(* IEC 61131-3 sources: kns-pump-station/src/POUs/Station/FB_LevelControlPid, 2 files *)

(* ---- FB_LevelControlPid.decl.st ---- *)
// Назначение: поддержание уровня ПИД LIC101 — число насосов и подключение подпорного по нагрузке
//             (04 §7.2), готовность ПИД (04 §7.4) с выдержкой STN_PID_RECOVER после восстановления
//             связи с ПЧ (04 §12), слежение ПИД за заданием ведущего, когда ПИД не управляет (04 §7.3);
//             выбыл ведущий при выбранном ПИД — выход держится (04 §7.3, §9).
//             Задание ПИД ФБ не считает: оно внешнее (stCfgLkg.rLevelSp_m, PRG_Station).
// Автор:      kr0nsch
// Версия:     0.2.1
// Документ:   docs/DESIGN.md, раздел 6.4; docs/04_algorithms.md, разделы 7, 12
FUNCTION_BLOCK FB_LevelControlPid
VAR_INPUT
    xEnable     : BOOL;             // eControlAct = LevelPid
    rLevel_m    : REAL;
    xLevelValid : BOOL;
    rPidOut_pct : REAL;             // GVL_Station.fbLIC101.rOut_pct (прошлый цикл)
    ePidMode    : PL.E_DeviceMode;  // GVL_Station.fbLIC101.Mode
    aitfPump    : ARRAY[1..GVL_Const.STN_PUMP_COUNT] OF PL.I_MotorVfd;
    axCommOk    : ARRAY[1..GVL_Const.STN_PUMP_COUNT] OF BOOL;   // нет MOT_WRN_COMM_LOSS
    uiLead      : UINT;             // ведущий (FB_PumpRotation, прошлый цикл); 0 — нет
    xInit       : BOOL;
    uiInitPumps : UINT;
    xPowerRestore : BOOL;           // нет напряжения или последовательный пуск (FB_PowerRestore): ПЧ без питания
                                    // или загружаются — нет связи, но это не потеря связи (VFD-12)
    itfTime     : PL.I_TimeSource;
END_VAR
VAR_IN_OUT CONSTANT
    stCfg : ST_StationCfg;          // rLvlStop_m, rLvlStartLead_m, rLvlStartAssist_m, tLvlConfirm,
                                    // rAssistOn_pct, tAssistOn, rAssistOff_pct, tAssistOff, uiDutyMax
END_VAR
VAR_OUTPUT
    uiRequired   : UINT;
    xPidReady    : BOOL;            // 04 §7.4; после восстановления связи — через STN_PID_RECOVER
    xPidControls : BOOL;            // xEnable AND ведущий SpeedAutoActive AND связь ведущего есть
    xTrack       : BOOL;            // → fbLIC101.xTrack (= NOT xPidControls)
    rTrack_pct   : REAL;            // → fbLIC101.rTrack_pct и rOutAct_pct: SpeedRef ведущего (0 — нет); ведущий
                                    // выбыл (Available = FALSE) при xEnable — rPidOut_pct: выход держится
END_VAR
VAR
    uiPumps        : UINT;          // состояние: 0, 1, 2 насоса
    fbStartLead    : PL.FB_Delay;   // 0 → 1: уровень >= rLvlStartLead_m (tLvlConfirm)
    fbAssistOnOut  : PL.FB_Delay;   // 1 → 2: выход ПИД >= rAssistOn_pct (tAssistOn)
    fbAssistOnLvl  : PL.FB_Delay;   // 1 → 2: уровень >= rLvlStartAssist_m (tLvlConfirm)
    fbAssistOff    : PL.FB_Delay;   // 2 → 1: выход ПИД <= rAssistOff_pct и уровень < rLvlStartAssist_m (tAssistOff)
    fbStopAll      : PL.FB_Delay;   // 1, 2 → 0: уровень <= rLvlStop_m (tLvlConfirm)
    fbCommRecover  : PL.FB_Delay;   // насос со связью есть: снятие сразу, возврат через STN_PID_RECOVER
    xFirstCall     : BOOL := TRUE;  // первый вызов: связь без выдержки возврата
END_VAR
VAR_TEMP
    uiMax          : UINT;          // MIN(STN_DUTY_MAX, uiDutyMax)
    uiPump         : UINT;          // номер насоса
    xAnyRunning    : BOOL;          // работает насос в Auto
    xCommRunning   : BOOL;          // работает насос в Auto со связью
    xCommAvailable : BOOL;          // доступен насос со связью (когда насосы стоят)
    xAnyAvailable  : BOOL;          // доступен хотя бы один насос
    xLeadValid     : BOOL;          // номер ведущего 1…STN_PUMP_COUNT и интерфейс задан
    xCommPart      : BOOL;          // есть насос со связью (условие готовности по связи)
    xCommBlock     : BOOL;          // насосы есть, но связи нет ни у одного: потеря связи
END_VAR

(* ---- FB_LevelControlPid.impl.st ---- *)
// Способ ПИД — не больше двух насосов (ведущий и подпорный) и не больше uiDutyMax
uiMax := MIN(GVL_Const.STN_DUTY_MAX, stCfg.uiDutyMax);
xLeadValid := uiLead >= 1 AND uiLead <= GVL_Const.STN_PUMP_COUNT;
IF xLeadValid THEN
    xLeadValid := aitfPump[uiLead] <> 0;
END_IF

// 1. Слежение (04 §7.3): ПИД управляет, только когда выбран, а ведущий работает в Auto без отказа
//    (SpeedAutoActive) и со связью с ПЧ; иначе выход следует за заданием ведущего (0 — ведущего нет).
//    Ведущий — прошлого цикла: если он выбыл (авария ПЧ, блокировка станции, смена режима — Available = FALSE),
//    роль в этом цикле передаст FB_PumpRotation, а остальные насосы работают с прежним заданием. Задание
//    выбывшего ПЧ (0) — не задание станции: при выбранном ПИД выход держится (04 §7.3, §9)
xPidControls := FALSE;
rTrack_pct := 0.0;
IF xLeadValid THEN
    rTrack_pct := aitfPump[uiLead].SpeedRef;
    xPidControls := xEnable AND aitfPump[uiLead].SpeedAutoActive AND axCommOk[uiLead];
    IF xEnable AND NOT aitfPump[uiLead].Available THEN
        rTrack_pct := rPidOut_pct;
    END_IF
END_IF
xTrack := NOT xPidControls;

// 2. Готовность (04 §7.4): ПИД в Auto, уровень годен и есть насос со связью — среди работающих в
//    Auto, а если насосы стоят — среди доступных. Если насосы есть, но связи нет ни у одного, —
//    потеря связи: готовность снимается сразу и возвращается через STN_PID_RECOVER (04 §12). Пока нет
//    напряжения или идёт последовательный пуск, ПЧ без питания или загружаются (VFD-12): связи нет, но это не
//    потеря — выдержка возврата не перезапускается, готовность — как только связь есть (04 §7.4)
xAnyRunning := FALSE;
xCommRunning := FALSE;
xCommAvailable := FALSE;
xAnyAvailable := FALSE;
FOR uiPump := 1 TO GVL_Const.STN_PUMP_COUNT DO
    IF aitfPump[uiPump] <> 0 THEN
        IF aitfPump[uiPump].Running AND aitfPump[uiPump].Mode = PL.E_DeviceMode.Auto THEN
            xAnyRunning := TRUE;
            xCommRunning := xCommRunning OR axCommOk[uiPump];
        END_IF
        IF aitfPump[uiPump].Available THEN
            xAnyAvailable := TRUE;
            xCommAvailable := xCommAvailable OR axCommOk[uiPump];
        END_IF
    END_IF
END_FOR
xCommPart := SEL(xAnyRunning, xCommAvailable, xCommRunning);
xCommBlock := SEL(xAnyRunning, xAnyAvailable, TRUE) AND NOT xCommPart;
IF xFirstCall THEN
    fbCommRecover.Preset(xValue := TRUE);           // при старте выдержки возврата нет
END_IF
fbCommRecover(xIn := NOT xCommBlock OR xPowerRestore, tOnDelay := GVL_Const.STN_PID_RECOVER, itfTime := itfTime);
xPidReady := ePidMode = PL.E_DeviceMode.Auto AND xLevelValid AND xCommPart AND fbCommRecover.xOut;

// 3. Вход без рывка: число насосов — по работающим, выдержки — заново
IF xInit THEN
    uiPumps := MIN(uiInitPumps, uiMax);
    fbStartLead.Preset(xValue := FALSE);
    fbAssistOnOut.Preset(xValue := FALSE);
    fbAssistOnLvl.Preset(xValue := FALSE);
    fbAssistOff.Preset(xValue := FALSE);
    fbStopAll.Preset(xValue := FALSE);
END_IF
uiPumps := MIN(uiPumps, uiMax);

// 4. Число насосов (таблица 04 §7.2). Условия по выходу ПИД — только когда ПИД управляет: выход
//    в слежении повторяет задание ведущего и о нагрузке не говорит. Недостоверный уровень —
//    условий по уровню нет, состояние держится
fbStartLead(xIn := xLevelValid AND uiPumps = 0 AND uiMax > 0 AND rLevel_m >= stCfg.rLvlStartLead_m,
            tOnDelay := stCfg.tLvlConfirm, itfTime := itfTime);
fbAssistOnOut(xIn := xPidControls AND uiPumps = 1 AND uiMax > 1 AND rPidOut_pct >= stCfg.rAssistOn_pct,
              tOnDelay := stCfg.tAssistOn, itfTime := itfTime);
fbAssistOnLvl(xIn := xLevelValid AND uiPumps = 1 AND uiMax > 1 AND rLevel_m >= stCfg.rLvlStartAssist_m,
              tOnDelay := stCfg.tLvlConfirm, itfTime := itfTime);
fbAssistOff(xIn := xPidControls AND uiPumps = 2 AND rPidOut_pct <= stCfg.rAssistOff_pct
                   AND xLevelValid AND rLevel_m < stCfg.rLvlStartAssist_m,
            tOnDelay := stCfg.tAssistOff, itfTime := itfTime);
fbStopAll(xIn := xLevelValid AND uiPumps > 0 AND rLevel_m <= stCfg.rLvlStop_m,
          tOnDelay := stCfg.tLvlConfirm, itfTime := itfTime);

IF fbStopAll.xOut THEN
    uiPumps := 0;
ELSIF fbAssistOff.xOut THEN
    uiPumps := 1;
ELSIF fbAssistOnOut.xOut OR fbAssistOnLvl.xOut THEN
    uiPumps := 2;
ELSIF fbStartLead.xOut THEN
    uiPumps := 1;
END_IF

uiRequired := SEL(xEnable, 0, uiPumps);
xFirstCall := FALSE;
